Fanuc KAREL source: KA00142.KL

PROGRAM KA00142
%NOLOCKGROUP
VAR
  SRC: ARRAY[2] OF SHORT
  DST: CONFIG
BEGIN
  SRC[1] = 2
  DST = SRC[1]
END KA00142
